{attribute 'linkalways'} 
{attribute 'no_explicit_call' := 'This FB is a CLASS and must be accessed using methods or properties'}
{attribute 'enable_dynamic_creation'}
FUNCTION_BLOCK _ETcVnSolvePnPMethod EXTENDS EnumDatatypeBase
VAR
	localData : ETcVnSolvePnPMethod;
	activeData : REFERENCE TO ETcVnSolvePnPMethod;
	enumBaseDatatype : _DINT(localData);
END_VAR

METHOD PRIVATE AddLocalEnumeration
VAR_INPUT
	Enumeration : T_MAXSTRING;
	Value : ETcVnSolvePnPMethod;
END_VAR
AddEnumeration(Enumeration, Value);
END_METHOD

PROPERTY PUBLIC Address : PVOID
GET
Address := ADR(activeData);
END_GET
END_PROPERTY

METHOD PUBLIC ClearReference
VAR_INPUT
END_VAR
activeData REF= localData;
SetBaseDatatypeReference();
END_METHOD

METHOD PUBLIC Clone : I_Datatype
VAR
    pClone : POINTER TO _ETcVnSolvePnPMethod;
END_VAR
pClone := __NEW(_ETcVnSolvePnPMethod(InitialValue := Value));
Clone := pClone^;
END_METHOD

METHOD FB_init : BOOL
VAR_INPUT
	bInitRetains : BOOL; // if TRUE, the retain variables are initialized (warm start / cold start)
	bInCopyCode : BOOL;  // if TRUE, the instance afterwards gets moved into the copy code (online change)
	InitialValue : ETcVnSolvePnPMethod;
END_VAR
localData := InitialValue;
AddBaseDatatype(enumBaseDatatype);
ClearReference();

AddLocalEnumeration('TCVN_SPM_ITERATIVE', ETcVnSolvePnPMethod.TCVN_SPM_ITERATIVE);
AddLocalEnumeration('TCVN_SPM_EPNP', ETcVnSolvePnPMethod.TCVN_SPM_EPNP);
AddLocalEnumeration('TCVN_SPM_P3P', ETcVnSolvePnPMethod.TCVN_SPM_P3P);
AddLocalEnumeration('TCVN_SPM_AP3P', ETcVnSolvePnPMethod.TCVN_SPM_AP3P);
AddLocalEnumeration('TCVN_SPM_IPPE', ETcVnSolvePnPMethod.TCVN_SPM_IPPE);
AddLocalEnumeration('TCVN_SPM_IPPE_SQUARE', ETcVnSolvePnPMethod.TCVN_SPM_IPPE_SQUARE);
AddLocalEnumeration('TCVN_SPM_SQPNP', ETcVnSolvePnPMethod.TCVN_SPM_SQPNP);
END_METHOD

PROPERTY PUBLIC Identifier : T_MAXSTRING
GET
Identifier := 'ETcVnSolvePnPMethod';
END_GET
END_PROPERTY

METHOD IsEnumeratorValueEqual : BOOL
VAR_INPUT
	Enumerator : I_KeyValueForwardEnumerator;
END_VAR
VAR
	storedValue : ETcVnSolvePnPMethod;
END_VAR
IF NOT Enumerator.TryGet(storedValue) THEN
	RETURN;
END_IF

IsEnumeratorValueEqual := storedValue = activeData;
END_METHOD

METHOD PUBLIC MakeReferenceTo
VAR_INPUT
	ReferenceTarget : REFERENCE TO ETcVnSolvePnPMethod;
END_VAR
activeData REF= ReferenceTarget;
SetBaseDatatypeReference();
END_METHOD

METHOD PROTECTED SetBaseDatatypeReference
VAR_INPUT
END_VAR
enumBaseDatatype.MakeReferenceTo(activeData);
END_METHOD

PROPERTY PUBLIC Size : UDINT
GET
Size := SIZEOF(activeData);
END_GET
END_PROPERTY

METHOD TryMakeReferenceTo : BOOL
VAR_INPUT
	Target : I_Datatype;
END_VAR
VAR
	pTargetData : POINTER TO ETcVnSolvePnPMethod;
END_VAR
IF NOT IsEquivalentTo(Target) THEN
	RETURN;
END_IF

pTargetData := Target.Address;
activeData REF= pTargetData^;
SetBaseDatatypeReference();
TryMakeReferenceTo := TRUE;
END_METHOD

PROPERTY PUBLIC Value : ETcVnSolvePnPMethod
GET
Value := activeData;
END_GET
SET
activeData := Value;
END_SET
END_PROPERTY

END_FUNCTION_BLOCK

(* stored: Version 1.1.0.1, ProductVersion 3.1.4024.13
   POU _ETcVnSolvePnPMethod: Id {93e8093c-f0d3-0ae1-1c04-9acab1a62f3b}, SpecialFunc None
   Folder Core: Id {c19d6535-904d-0fe6-2b2e-aa58d08509b6}
   Folder Protected: Id {d2569fe9-3811-0cb2-2fa6-bd3237163762}
   Folder Customize: Id {b5e5d6b6-5f53-003a-3e02-973acf7eaf9e}
   Folder Constructor: Id {e1e72cd6-2121-0341-3a12-482c02a9bec6}
   Folder Private: Id {0d7004be-713a-016e-12e9-06370cbd39a0}
   Folder Protected: Id {a9b2e5fb-7f96-04e7-2b6e-2ec8fcc537cf}
   Method AddLocalEnumeration: Id {7189cee1-cf8c-0819-1788-41e6672bbdfa}
   Property Address: Id {eba46181-4079-0009-226b-586f828059dc}
   Get Get: Id {6eb86ba4-97a6-061f-24fc-43a6e04e7462}
   Method ClearReference: Id {67887f0c-ccb1-0a97-2740-2c73f1526b33}
   Method Clone: Id {321b22b2-fd82-0fa7-2ed0-d75bb22d13d4}
   Method FB_init: Id {1bbb8533-c197-0d09-0b73-b8470fea1c8c}
   Property Identifier: Id {4a34e66d-68ec-0440-31bb-73f0b169bf20}
   Get Get: Id {740fbe4c-3d47-0c4a-03ba-938b2dcef0af}
   Method IsEnumeratorValueEqual: Id {e3e44a9e-0bec-09b5-212b-09a2c1514c5f}
   Method MakeReferenceTo: Id {42533c2a-89a9-09ce-08a5-4b97ea228537}
   Method SetBaseDatatypeReference: Id {fd8b2ca2-d6ef-0348-18ac-7982cbc912fa}
   Property Size: Id {71545f28-3044-0394-1060-3d028172f925}
   Get Get: Id {0aaef6d1-2a89-0024-22a6-8227bb27fdd0}
   Method TryMakeReferenceTo: Id {4ac1763b-39ce-0726-26fc-510432fb6ccc}
   Property Value: Id {258044b2-c23a-0509-2688-7c17eac4834c}
   Get Get: Id {229e6db7-a840-0490-19c5-33246ca5e40e}
   Set Set: Id {f7440bb4-bec9-0b62-3002-3881b70c97ad} *)
